ABB RAPID module: LongProg_0.modx

%%%
  VERSION:1
  LANGUAGE:ENGLISH
%%%
MODULE MOD_Tmp1

	PROC Prg_Tmp1()

		ConfJ \On;
		ConfL \Off;
		! Program generated by RoboDK v6.0.7 for ABB IRB 120-3/0.6 on XX/XX/XXXX 18:00:00
		! Using nominal kinematics.
		MoveAbsJ [[0.000000,-10.000000,20.000000,0.000000,30.000000,0.000000],[9E+09,9E+09,9E+09,9E+09,9E+09,9E+09]],v500,z1,ToolS \WObj:=FrameS;

	ENDPROC

ENDMODULE
